(* IEC 61131-3 sources: plc-vscode/tests/st/all/trust-platform/crates/trust-runtime/tests/fixtures/oscat/core/src/08_arithmetics_with_double_precision, 1 file *)

(* ---- tests.st ---- *)
TEST_PROGRAM oscat_math_real2_helpers_behave
VAR
    Base : REAL2;
    Sum1 : REAL2;
    Sum2 : REAL2;
    Product : REAL2;
    Negative : REAL2;
    Absolute : REAL2;
END_VAR

Base := R2_SET(X := REAL#1.5);
ASSERT_NEAR(EXPECTED := REAL#1.5, ACTUAL := Base.RX, DELTA := REAL#0.0001);
ASSERT_NEAR(EXPECTED := REAL#0.0, ACTUAL := Base.R1, DELTA := REAL#0.0001);

Sum1 := R2_ADD(X := Base, Y := REAL#0.25);
ASSERT_NEAR(EXPECTED := REAL#1.75, ACTUAL := Sum1.RX, DELTA := REAL#0.0001);
ASSERT_NEAR(EXPECTED := REAL#0.0, ACTUAL := Sum1.R1, DELTA := REAL#0.0001);

Sum2 := R2_ADD2(X := Base, Y := R2_SET(X := REAL#2.0));
ASSERT_NEAR(EXPECTED := REAL#3.5, ACTUAL := Sum2.RX, DELTA := REAL#0.0001);
ASSERT_NEAR(EXPECTED := REAL#0.0, ACTUAL := Sum2.R1, DELTA := REAL#0.0001);

Product := R2_MUL(X := Base, Y := REAL#2.0);
ASSERT_NEAR(EXPECTED := REAL#3.0, ACTUAL := Product.RX, DELTA := REAL#0.0001);
ASSERT_NEAR(EXPECTED := REAL#0.0, ACTUAL := Product.R1, DELTA := REAL#0.0001);

Negative.RX := REAL#-1.5;
Negative.R1 := REAL#-0.25;
Absolute := R2_ABS(X := Negative);
ASSERT_NEAR(EXPECTED := REAL#1.5, ACTUAL := Absolute.RX, DELTA := REAL#0.0001);
ASSERT_NEAR(EXPECTED := REAL#0.25, ACTUAL := Absolute.R1, DELTA := REAL#0.0001);
END_TEST_PROGRAM
